(* IEC 61131-3 sources: rusty/tests/lit/cfc/blocks/fb_call, 2 files *)

(* ---- main.st ---- *)
FUNCTION main : DINT
    fb_call();
    fb_call();
    // CHECK: a = 2, b = 20
    printf('a = %d, b = %d$N', fb_call.outA, fb_call.outB);
END_FUNCTION

(* ---- counter.st ---- *)
FUNCTION_BLOCK counter
VAR_INPUT
    step : DINT;
END_VAR
VAR_OUTPUT
    total : DINT;
END_VAR
    total := total + step;
END_FUNCTION_BLOCK
